// TIA Portal V20 export
FUNCTION "alarmy" : Void   // FC100, LAD
{ S7_Optimized_Access := 'TRUE' }
// stored: AutoNumber false, SetENOAutomatically false
   VAR_OUTPUT
      fc_alarm_global : Bool;
      fc_wrong_global : Bool;
      fc_op_1_alrm : Bool;
      fc_op_1_wrong : Bool;
      fc_op_2_alrm : Bool;
      fc_op_2_wrong : Bool;
      fc_op_3_alrm : Bool;
      fc_op_3_wrong : Bool;
   END_VAR
   VAR_TEMP
      OP_1_E : Bool;
      OP_2_E : Bool;
      OP_3_E : Bool;
      OP_4_E : Bool;
      OP_5_E : Bool;
      OP_1_W : Bool;
      OP_2_W : Bool;
      OP_3_W : Bool;
      OP_4_W : Bool;
      OP_5_W : Bool;
   END_VAR
   VAR CONSTANT
      TIME_ERROR_BOR : Time := T#4S;
   END_VAR
BEGIN

REGION Network 1: op_1 alarmy proces
END_REGION

REGION Network 2: op_1_warning_proces
END_REGION

REGION Network 3: OP_1_ALARM
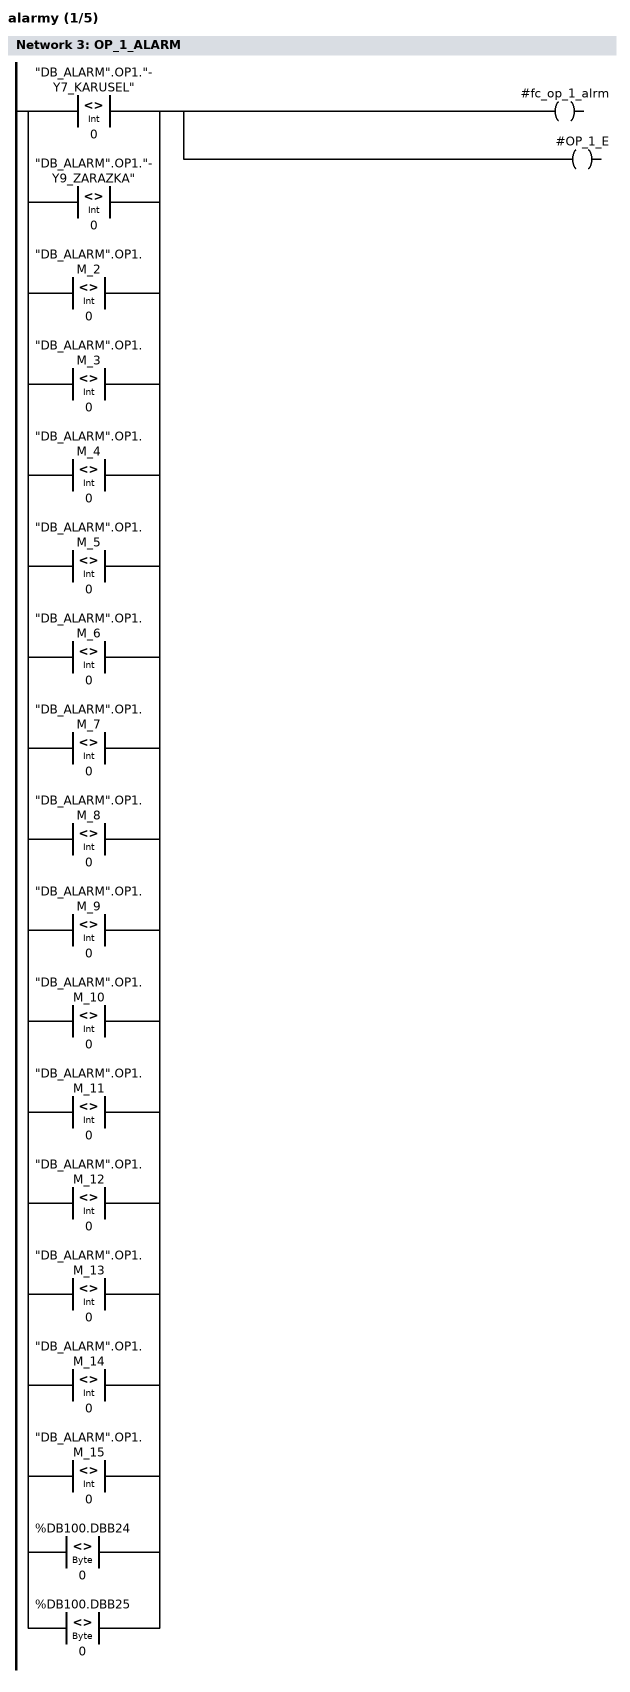
   RUNG wire#powerrail
      { S7_Templates := "SrcType := Int" } NE_Contact(in1 := "DB_ALARM".OP1."-Y7_KARUSEL", in2 := 0)
      wire#w1
      Coil( #fc_op_1_alrm )
   END_RUNG
   RUNG wire#powerrail
      { S7_Templates := "SrcType := Int" } NE_Contact(in1 := "DB_ALARM".OP1."-Y9_ZARAZKA", in2 := 0)
   END_RUNG wire#w1
   RUNG wire#powerrail
      { S7_Templates := "SrcType := Int" } NE_Contact(in1 := "DB_ALARM".OP1.M_2, in2 := 0)
   END_RUNG wire#w1
   RUNG wire#powerrail
      { S7_Templates := "SrcType := Int" } NE_Contact(in1 := "DB_ALARM".OP1.M_3, in2 := 0)
   END_RUNG wire#w1
   RUNG wire#powerrail
      { S7_Templates := "SrcType := Int" } NE_Contact(in1 := "DB_ALARM".OP1.M_4, in2 := 0)
   END_RUNG wire#w1
   RUNG wire#powerrail
      { S7_Templates := "SrcType := Int" } NE_Contact(in1 := "DB_ALARM".OP1.M_5, in2 := 0)
   END_RUNG wire#w1
   RUNG wire#powerrail
      { S7_Templates := "SrcType := Int" } NE_Contact(in1 := "DB_ALARM".OP1.M_6, in2 := 0)
   END_RUNG wire#w1
   RUNG wire#powerrail
      { S7_Templates := "SrcType := Int" } NE_Contact(in1 := "DB_ALARM".OP1.M_7, in2 := 0)
   END_RUNG wire#w1
   RUNG wire#powerrail
      { S7_Templates := "SrcType := Int" } NE_Contact(in1 := "DB_ALARM".OP1.M_8, in2 := 0)
   END_RUNG wire#w1
   RUNG wire#powerrail
      { S7_Templates := "SrcType := Int" } NE_Contact(in1 := "DB_ALARM".OP1.M_9, in2 := 0)
   END_RUNG wire#w1
   RUNG wire#powerrail
      { S7_Templates := "SrcType := Int" } NE_Contact(in1 := "DB_ALARM".OP1.M_10, in2 := 0)
   END_RUNG wire#w1
   RUNG wire#powerrail
      { S7_Templates := "SrcType := Int" } NE_Contact(in1 := "DB_ALARM".OP1.M_11, in2 := 0)
   END_RUNG wire#w1
   RUNG wire#powerrail
      { S7_Templates := "SrcType := Int" } NE_Contact(in1 := "DB_ALARM".OP1.M_12, in2 := 0)
   END_RUNG wire#w1
   RUNG wire#powerrail
      { S7_Templates := "SrcType := Int" } NE_Contact(in1 := "DB_ALARM".OP1.M_13, in2 := 0)
   END_RUNG wire#w1
   RUNG wire#powerrail
      { S7_Templates := "SrcType := Int" } NE_Contact(in1 := "DB_ALARM".OP1.M_14, in2 := 0)
   END_RUNG wire#w1
   RUNG wire#powerrail
      { S7_Templates := "SrcType := Int" } NE_Contact(in1 := "DB_ALARM".OP1.M_15, in2 := 0)
   END_RUNG wire#w1
   RUNG wire#powerrail
      { S7_Templates := "SrcType := Byte" } NE_Contact(in1 := %DB100.DBB24, in2 := 0)
   END_RUNG wire#w1
   RUNG wire#powerrail
      { S7_Templates := "SrcType := Byte" } NE_Contact(in1 := %DB100.DBB25, in2 := 0)
   END_RUNG wire#w1
   RUNG wire#w1
      Coil( #OP_1_E )
   END_RUNG
   // the same network as SCL:
   #fc_op_1_alrm := ("DB_ALARM".OP1."-Y7_KARUSEL" <> 0) OR ("DB_ALARM".OP1."-Y9_ZARAZKA" <> 0) OR ("DB_ALARM".OP1.M_2 <> 0) OR ("DB_ALARM".OP1.M_3 <> 0) OR ("DB_ALARM".OP1.M_4 <> 0) OR ("DB_ALARM".OP1.M_5 <> 0) OR ("DB_ALARM".OP1.M_6 <> 0) OR ("DB_ALARM".OP1.M_7 <> 0) OR ("DB_ALARM".OP1.M_8 <> 0) OR ("DB_ALARM".OP1.M_9 <> 0) OR ("DB_ALARM".OP1.M_10 <> 0) OR ("DB_ALARM".OP1.M_11 <> 0) OR ("DB_ALARM".OP1.M_12 <> 0) OR ("DB_ALARM".OP1.M_13 <> 0) OR ("DB_ALARM".OP1.M_14 <> 0) OR ("DB_ALARM".OP1.M_15 <> 0) OR (%DB100.DBB24 <> 0) OR (%DB100.DBB25 <> 0);
   #OP_1_E := #fc_op_1_alrm;
END_REGION

REGION Network 4: OP_2_ALARM
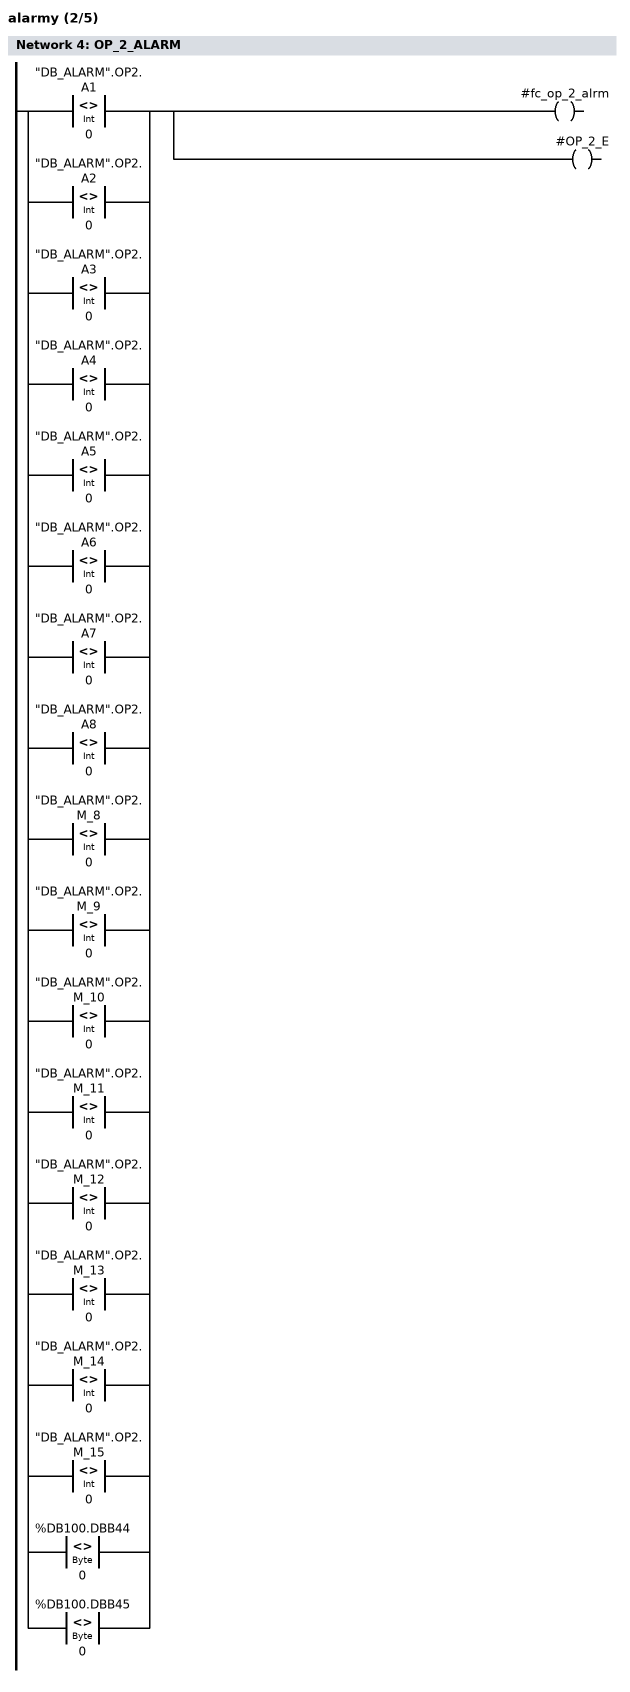
   RUNG wire#powerrail
      { S7_Templates := "SrcType := Int" } NE_Contact(in1 := "DB_ALARM".OP2.A1, in2 := 0)
      wire#w1
      Coil( #fc_op_2_alrm )
   END_RUNG
   RUNG wire#powerrail
      { S7_Templates := "SrcType := Int" } NE_Contact(in1 := "DB_ALARM".OP2.A2, in2 := 0)
   END_RUNG wire#w1
   RUNG wire#powerrail
      { S7_Templates := "SrcType := Int" } NE_Contact(in1 := "DB_ALARM".OP2.A3, in2 := 0)
   END_RUNG wire#w1
   RUNG wire#powerrail
      { S7_Templates := "SrcType := Int" } NE_Contact(in1 := "DB_ALARM".OP2.A4, in2 := 0)
   END_RUNG wire#w1
   RUNG wire#powerrail
      { S7_Templates := "SrcType := Int" } NE_Contact(in1 := "DB_ALARM".OP2.A5, in2 := 0)
   END_RUNG wire#w1
   RUNG wire#powerrail
      { S7_Templates := "SrcType := Int" } NE_Contact(in1 := "DB_ALARM".OP2.A6, in2 := 0)
   END_RUNG wire#w1
   RUNG wire#powerrail
      { S7_Templates := "SrcType := Int" } NE_Contact(in1 := "DB_ALARM".OP2.A7, in2 := 0)
   END_RUNG wire#w1
   RUNG wire#powerrail
      { S7_Templates := "SrcType := Int" } NE_Contact(in1 := "DB_ALARM".OP2.A8, in2 := 0)
   END_RUNG wire#w1
   RUNG wire#powerrail
      { S7_Templates := "SrcType := Int" } NE_Contact(in1 := "DB_ALARM".OP2.M_8, in2 := 0)
   END_RUNG wire#w1
   RUNG wire#powerrail
      { S7_Templates := "SrcType := Int" } NE_Contact(in1 := "DB_ALARM".OP2.M_9, in2 := 0)
   END_RUNG wire#w1
   RUNG wire#powerrail
      { S7_Templates := "SrcType := Int" } NE_Contact(in1 := "DB_ALARM".OP2.M_10, in2 := 0)
   END_RUNG wire#w1
   RUNG wire#powerrail
      { S7_Templates := "SrcType := Int" } NE_Contact(in1 := "DB_ALARM".OP2.M_11, in2 := 0)
   END_RUNG wire#w1
   RUNG wire#powerrail
      { S7_Templates := "SrcType := Int" } NE_Contact(in1 := "DB_ALARM".OP2.M_12, in2 := 0)
   END_RUNG wire#w1
   RUNG wire#powerrail
      { S7_Templates := "SrcType := Int" } NE_Contact(in1 := "DB_ALARM".OP2.M_13, in2 := 0)
   END_RUNG wire#w1
   RUNG wire#powerrail
      { S7_Templates := "SrcType := Int" } NE_Contact(in1 := "DB_ALARM".OP2.M_14, in2 := 0)
   END_RUNG wire#w1
   RUNG wire#powerrail
      { S7_Templates := "SrcType := Int" } NE_Contact(in1 := "DB_ALARM".OP2.M_15, in2 := 0)
   END_RUNG wire#w1
   RUNG wire#powerrail
      { S7_Templates := "SrcType := Byte" } NE_Contact(in1 := %DB100.DBB44, in2 := 0)
   END_RUNG wire#w1
   RUNG wire#powerrail
      { S7_Templates := "SrcType := Byte" } NE_Contact(in1 := %DB100.DBB45, in2 := 0)
   END_RUNG wire#w1
   RUNG wire#w1
      Coil( #OP_2_E )
   END_RUNG
   // the same network as SCL:
   #fc_op_2_alrm := ("DB_ALARM".OP2.A1 <> 0) OR ("DB_ALARM".OP2.A2 <> 0) OR ("DB_ALARM".OP2.A3 <> 0) OR ("DB_ALARM".OP2.A4 <> 0) OR ("DB_ALARM".OP2.A5 <> 0) OR ("DB_ALARM".OP2.A6 <> 0) OR ("DB_ALARM".OP2.A7 <> 0) OR ("DB_ALARM".OP2.A8 <> 0) OR ("DB_ALARM".OP2.M_8 <> 0) OR ("DB_ALARM".OP2.M_9 <> 0) OR ("DB_ALARM".OP2.M_10 <> 0) OR ("DB_ALARM".OP2.M_11 <> 0) OR ("DB_ALARM".OP2.M_12 <> 0) OR ("DB_ALARM".OP2.M_13 <> 0) OR ("DB_ALARM".OP2.M_14 <> 0) OR ("DB_ALARM".OP2.M_15 <> 0) OR (%DB100.DBB44 <> 0) OR (%DB100.DBB45 <> 0);
   #OP_2_E := #fc_op_2_alrm;
END_REGION

REGION Network 5: OP_3_ALARM
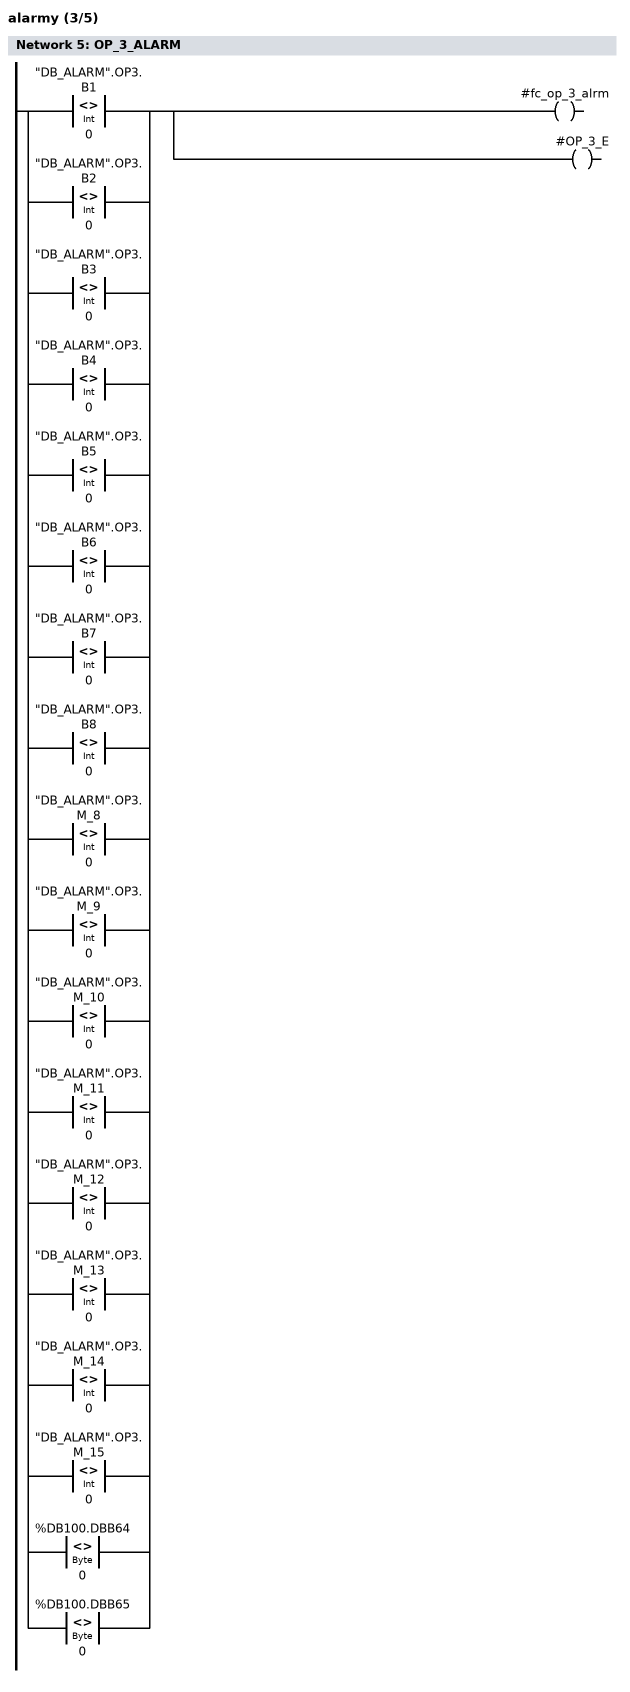
   RUNG wire#powerrail
      { S7_Templates := "SrcType := Int" } NE_Contact(in1 := "DB_ALARM".OP3.B1, in2 := 0)
      wire#w1
      Coil( #fc_op_3_alrm )
   END_RUNG
   RUNG wire#powerrail
      { S7_Templates := "SrcType := Int" } NE_Contact(in1 := "DB_ALARM".OP3.B2, in2 := 0)
   END_RUNG wire#w1
   RUNG wire#powerrail
      { S7_Templates := "SrcType := Int" } NE_Contact(in1 := "DB_ALARM".OP3.B3, in2 := 0)
   END_RUNG wire#w1
   RUNG wire#powerrail
      { S7_Templates := "SrcType := Int" } NE_Contact(in1 := "DB_ALARM".OP3.B4, in2 := 0)
   END_RUNG wire#w1
   RUNG wire#powerrail
      { S7_Templates := "SrcType := Int" } NE_Contact(in1 := "DB_ALARM".OP3.B5, in2 := 0)
   END_RUNG wire#w1
   RUNG wire#powerrail
      { S7_Templates := "SrcType := Int" } NE_Contact(in1 := "DB_ALARM".OP3.B6, in2 := 0)
   END_RUNG wire#w1
   RUNG wire#powerrail
      { S7_Templates := "SrcType := Int" } NE_Contact(in1 := "DB_ALARM".OP3.B7, in2 := 0)
   END_RUNG wire#w1
   RUNG wire#powerrail
      { S7_Templates := "SrcType := Int" } NE_Contact(in1 := "DB_ALARM".OP3.B8, in2 := 0)
   END_RUNG wire#w1
   RUNG wire#powerrail
      { S7_Templates := "SrcType := Int" } NE_Contact(in1 := "DB_ALARM".OP3.M_8, in2 := 0)
   END_RUNG wire#w1
   RUNG wire#powerrail
      { S7_Templates := "SrcType := Int" } NE_Contact(in1 := "DB_ALARM".OP3.M_9, in2 := 0)
   END_RUNG wire#w1
   RUNG wire#powerrail
      { S7_Templates := "SrcType := Int" } NE_Contact(in1 := "DB_ALARM".OP3.M_10, in2 := 0)
   END_RUNG wire#w1
   RUNG wire#powerrail
      { S7_Templates := "SrcType := Int" } NE_Contact(in1 := "DB_ALARM".OP3.M_11, in2 := 0)
   END_RUNG wire#w1
   RUNG wire#powerrail
      { S7_Templates := "SrcType := Int" } NE_Contact(in1 := "DB_ALARM".OP3.M_12, in2 := 0)
   END_RUNG wire#w1
   RUNG wire#powerrail
      { S7_Templates := "SrcType := Int" } NE_Contact(in1 := "DB_ALARM".OP3.M_13, in2 := 0)
   END_RUNG wire#w1
   RUNG wire#powerrail
      { S7_Templates := "SrcType := Int" } NE_Contact(in1 := "DB_ALARM".OP3.M_14, in2 := 0)
   END_RUNG wire#w1
   RUNG wire#powerrail
      { S7_Templates := "SrcType := Int" } NE_Contact(in1 := "DB_ALARM".OP3.M_15, in2 := 0)
   END_RUNG wire#w1
   RUNG wire#powerrail
      { S7_Templates := "SrcType := Byte" } NE_Contact(in1 := %DB100.DBB64, in2 := 0)
   END_RUNG wire#w1
   RUNG wire#powerrail
      { S7_Templates := "SrcType := Byte" } NE_Contact(in1 := %DB100.DBB65, in2 := 0)
   END_RUNG wire#w1
   RUNG wire#w1
      Coil( #OP_3_E )
   END_RUNG
   // the same network as SCL:
   #fc_op_3_alrm := ("DB_ALARM".OP3.B1 <> 0) OR ("DB_ALARM".OP3.B2 <> 0) OR ("DB_ALARM".OP3.B3 <> 0) OR ("DB_ALARM".OP3.B4 <> 0) OR ("DB_ALARM".OP3.B5 <> 0) OR ("DB_ALARM".OP3.B6 <> 0) OR ("DB_ALARM".OP3.B7 <> 0) OR ("DB_ALARM".OP3.B8 <> 0) OR ("DB_ALARM".OP3.M_8 <> 0) OR ("DB_ALARM".OP3.M_9 <> 0) OR ("DB_ALARM".OP3.M_10 <> 0) OR ("DB_ALARM".OP3.M_11 <> 0) OR ("DB_ALARM".OP3.M_12 <> 0) OR ("DB_ALARM".OP3.M_13 <> 0) OR ("DB_ALARM".OP3.M_14 <> 0) OR ("DB_ALARM".OP3.M_15 <> 0) OR (%DB100.DBB64 <> 0) OR (%DB100.DBB65 <> 0);
   #OP_3_E := #fc_op_3_alrm;
END_REGION

REGION Network 6: OP_1_WRONG
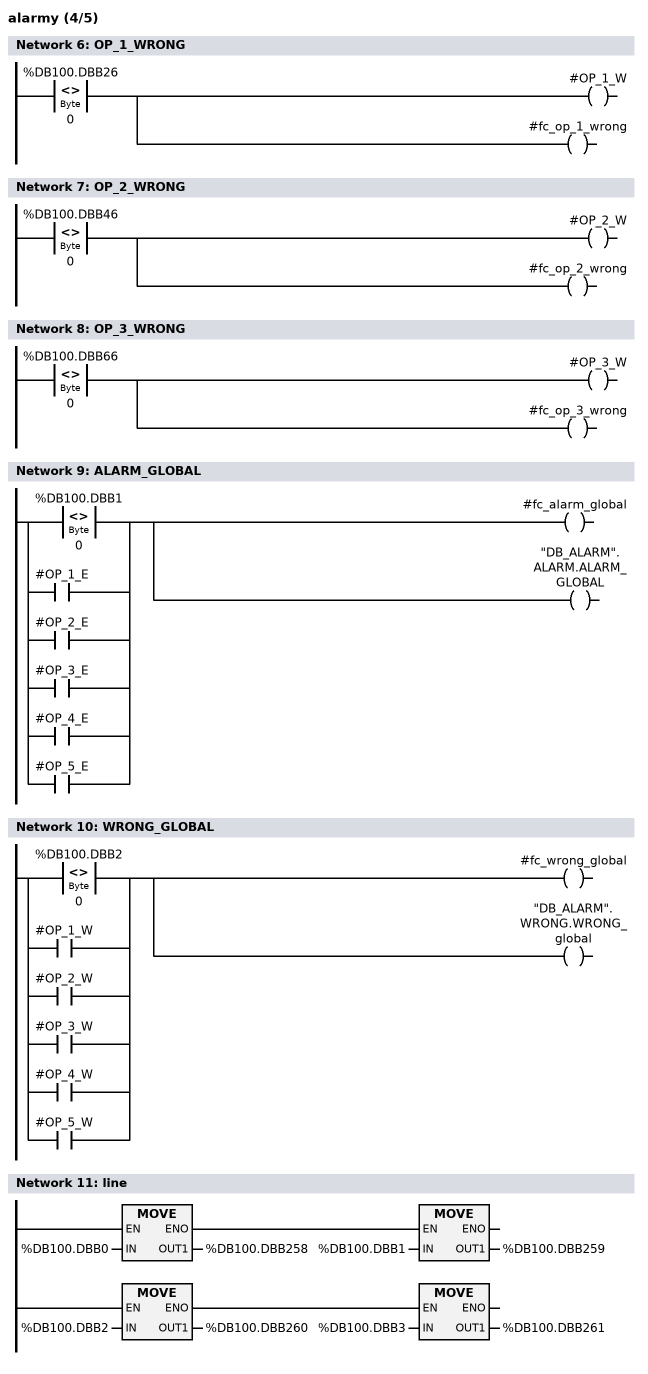
   RUNG wire#powerrail
      { S7_Templates := "SrcType := Byte" } NE_Contact(in1 := %DB100.DBB26, in2 := 0)
      wire#w1
      Coil( #OP_1_W )
   END_RUNG
   RUNG wire#w1
      Coil( #fc_op_1_wrong )
   END_RUNG
   // the same network as SCL:
   #OP_1_W := %DB100.DBB26 <> 0;
   #fc_op_1_wrong := #OP_1_W;
END_REGION

REGION Network 7: OP_2_WRONG
   RUNG wire#powerrail
      { S7_Templates := "SrcType := Byte" } NE_Contact(in1 := %DB100.DBB46, in2 := 0)
      wire#w1
      Coil( #OP_2_W )
   END_RUNG
   RUNG wire#w1
      Coil( #fc_op_2_wrong )
   END_RUNG
   // the same network as SCL:
   #OP_2_W := %DB100.DBB46 <> 0;
   #fc_op_2_wrong := #OP_2_W;
END_REGION

REGION Network 8: OP_3_WRONG
   RUNG wire#powerrail
      { S7_Templates := "SrcType := Byte" } NE_Contact(in1 := %DB100.DBB66, in2 := 0)
      wire#w1
      Coil( #OP_3_W )
   END_RUNG
   RUNG wire#w1
      Coil( #fc_op_3_wrong )
   END_RUNG
   // the same network as SCL:
   #OP_3_W := %DB100.DBB66 <> 0;
   #fc_op_3_wrong := #OP_3_W;
END_REGION

REGION Network 9: ALARM_GLOBAL
   RUNG wire#powerrail
      { S7_Templates := "SrcType := Byte" } NE_Contact(in1 := %DB100.DBB1, in2 := 0)
      wire#w1
      Coil( #fc_alarm_global )
   END_RUNG
   RUNG wire#powerrail
      Contact( #OP_1_E )
   END_RUNG wire#w1
   RUNG wire#powerrail
      Contact( #OP_2_E )
   END_RUNG wire#w1
   RUNG wire#powerrail
      Contact( #OP_3_E )
   END_RUNG wire#w1
   RUNG wire#powerrail
      Contact( #OP_4_E )
   END_RUNG wire#w1
   RUNG wire#powerrail
      Contact( #OP_5_E )
   END_RUNG wire#w1
   RUNG wire#w1
      Coil( "DB_ALARM".ALARM.ALARM_GLOBAL )
   END_RUNG
   // the same network as SCL:
   #fc_alarm_global := (%DB100.DBB1 <> 0) OR #OP_1_E OR #OP_2_E OR #OP_3_E OR #OP_4_E OR #OP_5_E;
   "DB_ALARM".ALARM.ALARM_GLOBAL := #fc_alarm_global;
END_REGION

REGION Network 10: WRONG_GLOBAL
   RUNG wire#powerrail
      { S7_Templates := "SrcType := Byte" } NE_Contact(in1 := %DB100.DBB2, in2 := 0)
      wire#w1
      Coil( #fc_wrong_global )
   END_RUNG
   RUNG wire#powerrail
      Contact( #OP_1_W )
   END_RUNG wire#w1
   RUNG wire#powerrail
      Contact( #OP_2_W )
   END_RUNG wire#w1
   RUNG wire#powerrail
      Contact( #OP_3_W )
   END_RUNG wire#w1
   RUNG wire#powerrail
      Contact( #OP_4_W )
   END_RUNG wire#w1
   RUNG wire#powerrail
      Contact( #OP_5_W )
   END_RUNG wire#w1
   RUNG wire#w1
      Coil( "DB_ALARM".WRONG.WRONG_global )
   END_RUNG
   // the same network as SCL:
   #fc_wrong_global := (%DB100.DBB2 <> 0) OR #OP_1_W OR #OP_2_W OR #OP_3_W OR #OP_4_W OR #OP_5_W;
   "DB_ALARM".WRONG.WRONG_global := #fc_wrong_global;
END_REGION

REGION Network 11: line
   RUNG wire#powerrail
      Move(in := %DB100.DBB0, out1 => %DB100.DBB258)
      Move(in := %DB100.DBB1, out1 => %DB100.DBB259)
   END_RUNG
   RUNG wire#powerrail
      Move(in := %DB100.DBB2, out1 => %DB100.DBB260)
      Move(in := %DB100.DBB3, out1 => %DB100.DBB261)
   END_RUNG
   // the same network as SCL:
   %DB100.DBB258 := %DB100.DBB0;
   %DB100.DBB259 := %DB100.DBB1;
   %DB100.DBB260 := %DB100.DBB2;
   %DB100.DBB261 := %DB100.DBB3;
END_REGION

REGION Network 12: op_1
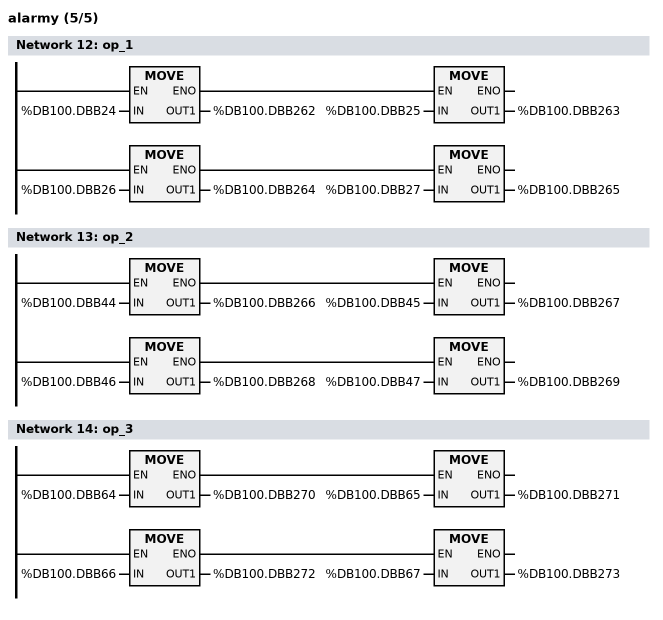
   RUNG wire#powerrail
      Move(in := %DB100.DBB24, out1 => %DB100.DBB262)
      Move(in := %DB100.DBB25, out1 => %DB100.DBB263)
   END_RUNG
   RUNG wire#powerrail
      Move(in := %DB100.DBB26, out1 => %DB100.DBB264)
      Move(in := %DB100.DBB27, out1 => %DB100.DBB265)
   END_RUNG
   // the same network as SCL:
   %DB100.DBB262 := %DB100.DBB24;
   %DB100.DBB263 := %DB100.DBB25;
   %DB100.DBB264 := %DB100.DBB26;
   %DB100.DBB265 := %DB100.DBB27;
END_REGION

REGION Network 13: op_2
   RUNG wire#powerrail
      Move(in := %DB100.DBB44, out1 => %DB100.DBB266)
      Move(in := %DB100.DBB45, out1 => %DB100.DBB267)
   END_RUNG
   RUNG wire#powerrail
      Move(in := %DB100.DBB46, out1 => %DB100.DBB268)
      Move(in := %DB100.DBB47, out1 => %DB100.DBB269)
   END_RUNG
   // the same network as SCL:
   %DB100.DBB266 := %DB100.DBB44;
   %DB100.DBB267 := %DB100.DBB45;
   %DB100.DBB268 := %DB100.DBB46;
   %DB100.DBB269 := %DB100.DBB47;
END_REGION

REGION Network 14: op_3
   RUNG wire#powerrail
      Move(in := %DB100.DBB64, out1 => %DB100.DBB270)
      Move(in := %DB100.DBB65, out1 => %DB100.DBB271)
   END_RUNG
   RUNG wire#powerrail
      Move(in := %DB100.DBB66, out1 => %DB100.DBB272)
      Move(in := %DB100.DBB67, out1 => %DB100.DBB273)
   END_RUNG
   // the same network as SCL:
   %DB100.DBB270 := %DB100.DBB64;
   %DB100.DBB271 := %DB100.DBB65;
   %DB100.DBB272 := %DB100.DBB66;
   %DB100.DBB273 := %DB100.DBB67;
END_REGION

REGION Network 15 (SCL)
   IF "CONTROL_LINE_DB".trig.reset_error_all = TRUE THEN
       // alarm global
       %DB100. := 0;
       %DB100. := 0;
       // wrong global
       %DB100. := 0;
       %DB100. := 0;
       // op_0
       // alarm
       %DB100. := 0;
       %DB100. := 0;
       // wrong
       %DB100. := 0;
       %DB100. := 0;
       // op_1
       // alarm
       %DB100. := 0;
       %DB100. := 0;
       // wrong
       %DB100. := 0;
       %DB100. := 0;
       // op_2
       // alarm
       %DB100. := 0;
       %DB100. := 0;
       // wrong
       %DB100. := 0;
       %DB100. := 0;
       // op_3
       // alarm
       %DB100. := 0;
       %DB100. := 0;
       // wrong
       %DB100. := 0;
       %DB100. := 0;
       // op_4
       // alarm
       %DB100. := 0;
       %DB100. := 0;
       // wrong
       %DB100. := 0;
       %DB100. := 0;
       // op_5
       // alarm
       %DB100. := 0;
       %DB100. := 0;
       // wrong
       %DB100. := 0;
       %DB100. := 0;
   END_IF;
END_REGION

REGION Network 16 (SCL)
   //"DB_ALARM".op_0_m_0 := "DB_ALARM".OP0.M_0;
   //"DB_ALARM".op_1_m_0 := "DB_ALARM".OP1.M_0;
   //"DB_ALARM".op_2_m_0 := "DB_ALARM".OP2.A1;
   //"DB_ALARM".op_2_m_1 := "DB_ALARM".OP2.A2;
   //"DB_ALARM".op_2_m_2 := "DB_ALARM".OP2.A3;
   //"DB_ALARM".op_2_m_3 := "DB_ALARM".OP2.A4;
   //"DB_ALARM".op_3_m_0 := "DB_ALARM".OP3.B1;
END_REGION
END_FUNCTION
